(* IEC 61131-3 sources: s7-to-codesys/s7conv/tests/snapshots/fixtures/src/POUs/FB_Broken, 1 file *)

(* ---- FB_Broken.decl.st ---- *)
// Назначение: Функциональный блок «FB_Broken», сконвертирован из SCL
// Автор:      не указан (исходный блок S7); перевод в ST — s7conv 0.1.0
// Версия:     0.1 (исходный блок S7)
// Документ:   docs/CONVERSION_REPORT.md, docs/MAPPING.md
// Источник:   s7conv/tests/fixtures/unsupported.scl, строки 46–53, FUNCTION_BLOCK "FB_Broken"
// Сгенерировано s7conv: пометки MIGRATION-CHECK и MIGRATION-TODO требуют ручного разбора.
FUNCTION_BLOCK FB_Broken
VAR_INPUT
    // MIGRATION-TODO: объявление не разобрано: ожидалось ';', найдено 'END_VAR' (стр. 49)
    // a : Int
END_VAR
